TYPE ST_GFX4IRTOPLC:
STRUCT
	nProcessVariable			:INT;
	wControllerStatus			:WORD;
	nOutputPower				:INT;
	wAmmeterInputOn			:WORD;
END_STRUCT
END_TYPE

(* stored: Version 1.1.0.1, ProductVersion 3.1.4024.15
   DUT ST_GFX4IRTOPLC: Id {e9db82c2-a89b-4375-bf8f-beec22a04c4d} *)
